FUNCTION F_time2seconds : REAL
VAR_INPUT
	tTime	:	TIME;
END_VAR
VAR
END_VAR

F_time2seconds	:=	TIME_TO_REAL(tTime) * CONVERSIONS.rTime2Seconds;

END_FUNCTION

(* stored: Version 1.1.0.1, ProductVersion 3.1.4024.9
   POU F_time2seconds: Id {8320d3a7-89fe-4fcd-accd-72e89d860407}, SpecialFunc None *)
